Fanuc KAREL source: KA00214.KL

PROGRAM KA00214
%NOLOCKGROUP
VAR
  SRC: ARRAY[4] OF XYZWPR
  DST: ARRAY[4] OF VECTOR
BEGIN
  DST = SRC
END KA00214
